// TIA Portal V20 export
DATA_BLOCK "T3_Datos"   // DB40939
{ S7_Optimized_Access := 'TRUE' }
AUTHOR : IA
FAMILY : PRUEBA
VERSION : 0.1
// Prueba IA 3: datos
// stored: AutoNumber false
   VAR
      Rama_1 : Bool;
      Rama_2 : Bool;
      Mul_Out : Int;
      Div_Out : Int;
      Ret_A : Int;
      Ret_B : Int;
   END_VAR
BEGIN
END_DATA_BLOCK
